(*
SPDX-FileCopyrightText: © 2026 Oleksandr Tiutyk <trofimich@gmail.com>
SPDX-License-Identifier: MIT
License: https://opensource.org/license/mit
*)

(*!
<summary>Provides fluent assertions on a copied LTIME value.</summary>
<description>
Copies actual into persistent instance storage before the entry method returns; literals and expression
results therefore remain valid throughout the immediate chain. Owns no heap allocation or pointed-to resource.
The message prefixes every failure until the next preparation. Finish one chain before starting another on
the owning Assertions provider. Use only from the owning test callback on one task, without reentry.
Obtain this context from the owning provider; direct unprepared use is unsupported.
Expected arguments use the declared IEC type; ordinary compiler conversions happen before comparison.
This context does not depend on another assertion context.
Object metadata is available before preparation; inherited equality compares instance identity.
</description>
*)

{attribute 'no_explicit_call' := 'do not call this function block directly'}
FUNCTION_BLOCK LongTimeAssertionContext EXTENDS TOF_Core.Object
VAR_STAT
	{attribute 'hide'}
	_ClassName : STRING := __POUNAME();
END_VAR
VAR
	_Actual : LTIME;
	_TestCase : ITestCase;
	_Message : WSTRING(255);
END_VAR

(*!
<summary>Provides the implementation class name.</summary>
<description>
Borrowed read-only reference to compiler-initialized storage, valid throughout the instance lifetime.
Do not modify the returned reference; no ownership is transferred.
</description>
*)
{attribute 'monitoring' := 'call'}
PROPERTY ClassName : REFERENCE TO STRING
GET
ClassName REF= _ClassName;
END_GET
END_PROPERTY

(*!
<summary>Asserts that the actual value is strictly greater than expected.</summary>
<description>
Records failure without interrupting the callback; preserves the message for the rest of the chain.
</description>
<param name="expected">Expected value converted by the compiler to LTIME.</param>
*)
METHOD FINAL IsGreaterThan : REFERENCE TO LongTimeAssertionContext
VAR_INPUT
	expected : LTIME;
END_VAR
IF _Actual <= expected THEN
	failComparison(
		expected := expected,
		expectation := "Expected value > "
	);
END_IF

IsGreaterThan REF= THIS^;
END_METHOD

(*!
<summary>Asserts that the actual value meets the inclusive lower boundary.</summary>
<description>
Records failure without interrupting the callback; preserves the message for the rest of the chain.
</description>
<param name="expected">Expected value converted by the compiler to LTIME.</param>
*)
METHOD FINAL IsGreaterThanOrEquals : REFERENCE TO LongTimeAssertionContext
VAR_INPUT
	expected : LTIME;
END_VAR
IF _Actual < expected THEN
	failComparison(
		expected := expected,
		expectation := "Expected value >= "
	);
END_IF

IsGreaterThanOrEquals REF= THIS^;
END_METHOD

(*!
<summary>Asserts that the actual value is strictly less than expected.</summary>
<description>
Records failure without interrupting the callback; preserves the message for the rest of the chain.
</description>
<param name="expected">Expected value converted by the compiler to LTIME.</param>
*)
METHOD FINAL IsLessThan : REFERENCE TO LongTimeAssertionContext
VAR_INPUT
	expected : LTIME;
END_VAR
IF _Actual >= expected THEN
	failComparison(
		expected := expected,
		expectation := "Expected value < "
	);
END_IF

IsLessThan REF= THIS^;
END_METHOD

(*!
<summary>Asserts that the actual value meets the inclusive upper boundary.</summary>
<description>
Records failure without interrupting the callback; preserves the message for the rest of the chain.
</description>
<param name="expected">Expected value converted by the compiler to LTIME.</param>
*)
METHOD FINAL IsLessThanOrEquals : REFERENCE TO LongTimeAssertionContext
VAR_INPUT
	expected : LTIME;
END_VAR
IF _Actual > expected THEN
	failComparison(
		expected := expected,
		expectation := "Expected value <= "
	);
END_IF

IsLessThanOrEquals REF= THIS^;
END_METHOD

(*!
<summary>Provides the library namespace.</summary>
<description>
Borrowed read-only reference to the compiler-initialized namespace, valid throughout the instance lifetime.
Do not modify the returned reference; no ownership is transferred.
</description>
*)
{attribute 'monitoring' := 'call'}
PROPERTY NamespaceName : REFERENCE TO STRING
GET
NamespaceName REF= CurrentNamespace.Name;
END_GET
END_PROPERTY

(*!
<summary>Asserts inequality with the expected value.</summary>
<description>
Records failure without interrupting the callback; preserves the message for the rest of the chain.
</description>
<param name="expected">Expected value converted by the compiler to LTIME.</param>
*)
METHOD FINAL NotToBe : REFERENCE TO LongTimeAssertionContext
VAR_INPUT
	expected : LTIME;
END_VAR
IF _Actual = expected THEN
	failComparison(
		expected := expected,
		expectation := "Expected value not to be: "
	);
END_IF

NotToBe REF= THIS^;
END_METHOD

(*!
<summary>Copies the actual operand and replaces the chain-wide message.</summary>
<description>
Called by the owning Assertions provider after it verifies the running test case.
No pointer to this method's input storage is retained. The receiver is borrowed until the next preparation;
the owning provider keeps it alive throughout the immediate chain.
</description>
<param name="actual">Value copied into this context.</param>
<param name="testCase">Borrowed failure receiver for the immediate chain.</param>
<param name="message">Copied diagnostic prefix, including empty to clear the previous prefix.</param>
*)
METHOD INTERNAL FINAL Prepare
VAR_INPUT
	actual : LTIME;
	testCase : ITestCase;
	message : WSTRING(255);
END_VAR
_Actual := actual;
_TestCase := testCase;
_Message := message;
END_METHOD

(*!
<summary>Reports the byte size of this concrete instance.</summary>
<description>
Includes inline fields and nested instances, but excludes separately allocated payloads.
Obtaining the size does not transfer ownership or validate an arbitrary address.
</description>
*)
{attribute 'monitoring' := 'call'}
PROPERTY SelfSize : ULINT
GET
SelfSize := XSIZEOF(THIS^);
END_GET
END_PROPERTY

(*!
<summary>Asserts equality with the expected value.</summary>
<description>
Records failure without interrupting the callback; preserves the message for the rest of the chain.
</description>
<param name="expected">Expected value converted by the compiler to LTIME.</param>
*)
METHOD FINAL ToBe : REFERENCE TO LongTimeAssertionContext
VAR_INPUT
	expected : LTIME;
END_VAR
IF _Actual <> expected THEN
	failComparison(
		expected := expected,
		expectation := "Expected: "
	);
END_IF

ToBe REF= THIS^;
END_METHOD

(*!
<summary>Formats a failed typed predicate and reports it with the chain message.</summary>
<description>
Does not change operands or chain state. The receiver retains its first failure. Reporting exceptions
propagate to the enclosing test callback handler; an unprepared receiver is a configuration error.
</description>
<param name="expected">Typed expected operand used only for this diagnostic.</param>
<param name="expectation">Prefix identifying the failed predicate.</param>
*)
METHOD PRIVATE failComparison
VAR_INPUT
	expected : LTIME;
	expectation : WSTRING(40);
END_VAR
VAR
	actualText : WSTRING(255);
	expectedText : WSTRING(255);
	diagnostic : TOF_Core.ERROR_MESSAGE;
END_VAR
actualText := TO_WSTRING(_Actual);
expectedText := TO_WSTRING(expected);

diagnostic := TOF_Core.WideStrings.Concat255(
	expectation,
	expectedText,
	", but was: ",
	actualText
);

TestServices.ReportAssertionFailure(
	testCase := _TestCase,
	message := _Message,
	sourceClassName := ClassName,
	defaultMessage := diagnostic
);
END_METHOD

END_FUNCTION_BLOCK

(* stored: Version 1.1.0.1
   POU LongTimeAssertionContext: Id {2c0f4aa6-3a38-4c40-941e-7a3487cab9cd}, SpecialFunc None
   Folder Service methods: Id {d497960b-2432-431f-aa90-a2ddf100e8ee}
   Property ClassName: Id {fdda2eb1-15fa-437d-ad5b-8edfaafa2e16}
   Get Get: Id {356b269f-0f65-4f87-9207-7e4e9b74cf3e}
   Method IsGreaterThan: Id {f43c1443-ddae-42ac-a621-22ee48fc4eb9}
   Method IsGreaterThanOrEquals: Id {0e8063e1-7b91-45eb-b39f-6a9d3c6555ed}
   Method IsLessThan: Id {febf0a30-5749-40aa-ac09-5ac34fa48951}
   Method IsLessThanOrEquals: Id {b5aca956-e58a-4aa0-869e-ee6383d6a7d2}
   Property NamespaceName: Id {28818bb7-d9fd-4758-bce8-4c32fc077e22}
   Get Get: Id {9d1e87d4-b634-431f-b8e6-52a3f33038ec}
   Method NotToBe: Id {1aaeb720-8953-4245-a646-4011e291b0dd}
   Method Prepare: Id {2507650b-34f1-444d-ad1e-9bd6c7f6d86f}
   Property SelfSize: Id {65d16249-55c5-45d6-91f4-5b68a6746993}
   Get Get: Id {900d8f88-569c-422a-8ea6-5ff9923ecb06}
   Method ToBe: Id {330db42f-8668-4fc9-bee0-12447587ee1c}
   Method failComparison: Id {70ae8c84-1b5b-4a79-8d34-bec7360c49a3} *)
